ABB RAPID module: Prog_Name_Tha.prg

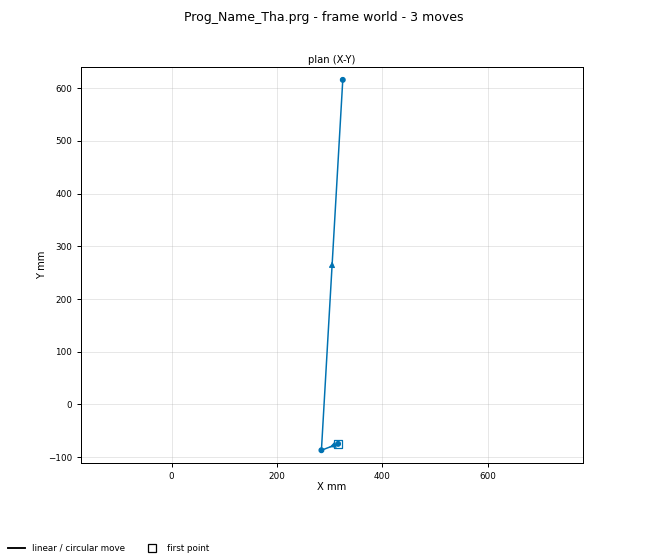
[picture p0: tool path of Prog_Name_Tha.prg in frame world, 3 of 5 moves have a stored position in this frame; points joined in program order, loops and branches not executed]
%%%
  VERSION:1
  LANGUAGE:ENGLISH
%%%
MODULE MOD_Prog_Name_Tha

    ! -------------------------------
    ! Define customized variables here
    ! ...

	! Tool variables:
	PERS tooldata Spindle := [TRUE,[[10.000,0.000,120.000],[0.99144486,0.00000000,0.13052619,0.00000001]],[1,[0,0,20],[1,0,0,0],0,0,0.005]];
	PERS tooldata Tool7 := [TRUE,[[10.000,0.000,120.000],[0.99144486,0.00000000,0.13052619,0.00000001]],[1,[0,0,20],[1,0,0,0],0,0,0.005]];

	! Reference variables:
	PERS wobjdata ABBIRB120306B := [FALSE, TRUE, "", [[0.000,0.000,0.000],[1.00000000,0.00000000,0.00000000,0.00000000]],[[0,0,0],[1,0,0,0]]];
	PERS wobjdata Frame12 := [FALSE, TRUE, "", [[250.000,300.000,-10.000],[0.70710678,0.00000000,0.00000000,0.70710678]],[[0,0,0],[1,0,0,0]]];

	PROC Main()
		ConfJ \On;
		ConfL \Off;
		! Program generated by VerticalBot Studio for ABB IRB 120-3/0.6 on 25/10/2026 12:00:00
		! Using nominal kinematics.
		MoveAbsJ [[-10.000000,10.000000,20.000000,30.000000,40.000000,-50.000000],[9E+09,9E+09,9E+09,9E+09,9E+09,9E+09]],v1000,z10,Spindle \WObj:=ABBIRB120306B;
		MoveL [[315.779,-74.668,245.881],[0.09884449,0.01379658,0.99324025,0.05927254],[-1,0,-1,0],[9E+09,9E+09,9E+09,9E+09,9E+09,9E+09]],v1000,z10,Spindle \WObj:=ABBIRB120306B;
		MoveL [[284.148,-86.783,243.844],[0.09359571,0.04936652,0.99254150,0.06053239],[-1,0,-1,0],[9E+09,9E+09,9E+09,9E+09,9E+09,9E+09]],v1000,[FALSE,0.5,0.8,0.8,0.1,0.8,0.1],Spindle \WObj:=ABBIRB120306B;
		STOP;
		WaitTime 1.500;
		TPWrite "Say "hi" to the operator";
		! A long comment line that exceeds the usual controller limits for comments by far, really
		SetDO D_OUT_12, 0;
		SetDO OUT_A, 1;
		WaitDI D_IN_4, 0, \MaxTime:=1.0;
		WaitDI IN_B, 1;
		Program_With_A_Long_Name_ABCDEFGHIJ;
		MoveL [[315.779,-74.668,245.881],[0.09884449,0.01379658,0.99324025,0.05927254],[-1,0,-1,0],[9E+09,9E+09,9E+09,9E+09,9E+09,9E+09]],v1000,[FALSE,0.5,0.8,0.8,0.1,0.8,0.1],Tool7 \WObj:=Frame12;
		MoveAbsJ [[-10.000000,10.000000,20.000000,30.000000,40.000000,-50.000000],[9E+09,9E+09,9E+09,9E+09,9E+09,9E+09]],v1000,fine,Tool7 \WObj:=Frame12;
	ENDPROC

ENDMODULE
